// TIA Portal V19 export
DATA_BLOCK "dummy"   // DB102
{ S7_Optimized_Access := 'FALSE' }
   VAR
      cheking_sp : Real;
      check_2 : Bool;
      check3 : Bool;
      R1 : Struct
         Intl_1 : Bool;
         Intl_2 : Bool;
         Intl_3 : Bool;
         Intl_4 : Bool;
      END_STRUCT;
      R2 : Struct
         Intl_1 : Bool;
         Intl_2 : Bool;
         Intl_3 : Bool;
         Intl_4 : Bool;
      END_STRUCT;
      R3 : Struct
         Intl_1 : Bool;
         Intl_2 : Bool;
         Intl_3 : Bool;
         Intl_4 : Bool;
      END_STRUCT;
      R4 : Struct
         Intl_1 : Bool;
         Intl_2 : Bool;
         Intl_3 : Bool;
         Intl_4 : Bool;
      END_STRUCT;
      R5 : Struct
         Intl_1 : Bool;
         Intl_2 : Bool;
         Intl_3 : Bool;
         Intl_4 : Bool;
      END_STRUCT;
      R6 : Struct
         Intl_1 : Bool;
         Intl_2 : Bool;
         Intl_3 : Bool;
         Intl_4 : Bool;
      END_STRUCT;
      R7 : Struct
         Intl_1 : Bool;
         Intl_2 : Bool;
         Intl_3 : Bool;
         Intl_4 : Bool;
      END_STRUCT;
      R8 : Struct
         Intl_1 : Bool;
         Intl_2 : Bool;
         Intl_3 : Bool;
         Intl_4 : Bool;
      END_STRUCT;
      R9 : Struct
         Intl_1 : Bool;
         Intl_2 : Bool;
         Intl_3 : Bool;
         Intl_4 : Bool;
      END_STRUCT;
      R10 : Struct
         Intl_1 : Bool;
         Intl_2 : Bool;
         Intl_3 : Bool;
         Intl_4 : Bool;
      END_STRUCT;
      R11 : Struct
         Intl_1 : Bool;
         Intl_2 : Bool;
         Intl_3 : Bool;
         Intl_4 : Bool;
      END_STRUCT;
      R12 : Struct
         Intl_1 : Bool;
         Intl_2 : Bool;
         Intl_3 : Bool;
         Intl_4 : Bool;
      END_STRUCT;
      R13 : Struct
         Intl_1 : Bool;
         Intl_2 : Bool;
         Intl_3 : Bool;
         Intl_4 : Bool;
      END_STRUCT;
      R14 : Struct
         Intl_1 : Bool;
         Intl_2 : Bool;
         Intl_3 : Bool;
         Intl_4 : Bool;
      END_STRUCT;
      R15 : Struct
         Intl_1 : Bool;
         Intl_2 : Bool;
         Intl_3 : Bool;
         Intl_4 : Bool;
      END_STRUCT;
      R16 : Struct
         Intl_1 : Bool;
         Intl_2 : Bool;
         Intl_3 : Bool;
         Intl_4 : Bool;
      END_STRUCT;
      R17 : Struct
         Intl_1 : Bool;
         Intl_2 : Bool;
         Intl_3 : Bool;
         Intl_4 : Bool;
      END_STRUCT;
      R18 : Struct
         Intl_1 : Bool;
         Intl_2 : Bool;
         Intl_3 : Bool;
         Intl_4 : Bool;
      END_STRUCT;
      SEMI_AUTO_SEL : Struct
         R1 : Int;
         R2 : Int;
         R3 : Int;
         R4 : Int;
         R5 : Int;
         R6 : Int;
         R7 : Int;
         R8 : Int;
         R9 : Int;
         R10 : Int;
         R11 : Int;
         R12 : Int;
         R13 : Int;
         R14 : Int;
         R15 : Int;
         R16 : Int;
         R17 : Int;
         R18 : Int;
      END_STRUCT;
      AG_STATUS : Struct
         R1 : Bool;
         R2 : Bool;
         R3 : Bool;
         R4 : Bool;
         R5 : Bool;
         R6 : Bool;
         R7 : Bool;
         R8 : Bool;
         R9 : Bool;
         R10 : Bool;
         R11 : Bool;
         R12 : Bool;
         R13 : Bool;
         R14 : Bool;
         R15 : Bool;
         R16 : Bool;
         R17 : Bool;
         R18 : Bool;
      END_STRUCT;
   END_VAR
BEGIN
END_DATA_BLOCK
